Staubli VAL3: insertSwitch.pgx

public program insertSwitch(string x_sKey, num x_nIndex, string x_sValue, bool x_bToSave)
  local num l_i
begin
  if x_nIndex==0 and progTemp:pProgItem[x_sKey].pProgTemplate[x_nIndex].sTRAJname==""
    x_nIndex=x_nIndex
  else
    x_nIndex=x_nIndex+1
    //insert(progTemp:pProgItem[x_sKey].pProgTemplate[x_nIndex])
    //l_nIndex=x_nIndex+1
    //insert(progTemp:pProgItem[x_sKey].pProgTemplate[x_nIndex+1])
    append(progTemp:pProgItem[x_sKey].pProgTemplate)
    for l_i = size(progTemp:pProgItem[x_sKey].pProgTemplate)-1 to x_nIndex step -1
      call copyPara(x_sKey,l_i-1,l_i)
    endFor
  endIf

  progTemp:pProgItem[x_sKey].pProgTemplate[x_nIndex].nType=5
  progTemp:pProgItem[x_sKey].pProgTemplate[x_nIndex].sTRAJname="SWITCH"
  progTemp:pProgItem[x_sKey].pProgTemplate[x_nIndex].sSwitchItem.sIOValue=x_sValue
  progTemp:pProgItem[x_sKey].pProgTemplate[x_nIndex].sSwitchItem.bIOdisable=true
  //insert(progTemp:pProgItem[x_sKey].pProgTemplate[x_nIndex+1])
  append(progTemp:pProgItem[x_sKey].pProgTemplate)
  for l_i = size(progTemp:pProgItem[x_sKey].pProgTemplate)-1 to(x_nIndex+1) step -1
    call copyPara(x_sKey,l_i-1,l_i)
  endFor
  progTemp:pProgItem[x_sKey].pProgTemplate[x_nIndex+1].nType=7
  progTemp:pProgItem[x_sKey].pProgTemplate[x_nIndex+1].sTRAJname="ENDSWITCH"
  //progTemp:pProgItem[x_sKey].pProgTemplate[x_nIndex].sSwitchItem.sIOValue=x_nValue
  //progTemp:pProgItem[x_sKey].pProgTemplate[x_nIndex].sSwitchItem.bIOdisable=true

  x_bToSave=true
end
